(*
SPDX-FileCopyrightText: © 2026 Oleksandr Tiutyk <trofimich@gmail.com>
SPDX-License-Identifier: MIT
License: https://opensource.org/license/mit
*)

(*!
<summary>Provides a scalar natural order for borrowed OBJECT list entries.</summary>
<description>
Supports other ICollectionSortValue objects. Comparisons copy the other scalar key without mutating or
retaining either object. The caller keeps sort keys stable during sorting; no allocation or cleanup is used.
</description>
*)

FUNCTION_BLOCK CollectionComparableProbe EXTENDS TOF_Core.Object IMPLEMENTS ICollectionSortValue
VAR_INPUT
	//! <summary>Scalar key defining the fixture's natural order.</summary>
	SortValue : DINT;
END_VAR
VAR_STAT
	_ClassName : STRING := __POUNAME();
END_VAR

(*!
<summary>Provides the concrete test fixture class name.</summary>
*)
{attribute 'monitoring' := 'call'}
PROPERTY ClassName : REFERENCE TO STRING
GET
ClassName REF= _ClassName;
END_GET
END_PROPERTY

(*!
<summary>Compares supported scalar-key objects and rejects null or unrelated comparable types.</summary>
*)
METHOD CompareTo : TOF_Core.COMPARISON_RESULT
VAR_IN_OUT CONSTANT
	otherValue : TOF_Core.IComparable;
END_VAR
VAR
	otherSortValue : ICollectionSortValue;
	otherKey : DINT;
END_VAR
IF otherValue = 0 THEN
	TOF_Core.Exceptions.ThrowArgumentNotSpecified(
		sourceNamespaceName := NamespaceName,
		sourceClassName := ClassName,
		sourcePOUName := __POUNAME(),
		sourcePosition := __POSITION(),
		argumentName := 'otherValue'
	);
END_IF

IF NOT __QUERYINTERFACE(otherValue, otherSortValue) THEN
	TOF_Core.Exceptions.ThrowStandard(
		sourceNamespaceName := NamespaceName,
		sourceClassName := ClassName,
		sourcePOUName := __POUNAME(),
		sourcePosition := __POSITION(),
		message := "Unsupported collection comparable fixture"
	);
END_IF

otherKey := otherSortValue.GetSortValue();

IF SortValue < otherKey THEN
	CompareTo := TOF_Core.COMPARISON_RESULT.FIRST_LESS_THAN_SECOND;
ELSIF SortValue > otherKey THEN
	CompareTo := TOF_Core.COMPARISON_RESULT.FIRST_GREATER_THAN_SECOND;
ELSE
	CompareTo := TOF_Core.COMPARISON_RESULT.FIRST_EQUAL_TO_SECOND;
END_IF
END_METHOD

(*!
<summary>Copies the configured sort key without mutation.</summary>
*)
METHOD GetSortValue : DINT
GetSortValue := SortValue;
END_METHOD

(*!
<summary>Borrows the compiler-initialized test namespace.</summary>
*)
{attribute 'monitoring' := 'call'}
PROPERTY NamespaceName : REFERENCE TO STRING
GET
NamespaceName REF= CurrentNamespace.Name;
END_GET
END_PROPERTY

(*!
<summary>Reports the complete fixture instance size, excluding separately allocated storage.</summary>
*)
{attribute 'monitoring' := 'call'}
PROPERTY SelfSize : ULINT
GET
SelfSize := XSIZEOF(THIS^);
END_GET
END_PROPERTY

END_FUNCTION_BLOCK

(* stored: Version 1.1.0.1, ProductVersion 3.1.4026.21
   POU CollectionComparableProbe: Id {be1ce13d-533b-447e-b1ca-bc68f369e23c}, SpecialFunc None
   Property ClassName: Id {524c25fa-effd-47d2-899c-109cd5d7359a}
   Get Get: Id {ff64f80e-ffa8-467f-b97b-1226aa0f4865}
   Method CompareTo: Id {ac7bfd62-7bdb-4ae7-a745-a4778e7bded0}
   Method GetSortValue: Id {356150dc-a1f2-4d5a-86ce-b5786a3643b8}
   Property NamespaceName: Id {362a1566-5de6-4e9b-a852-0a7ebe305c75}
   Get Get: Id {b0bab4ca-9949-451d-a46c-f9767d6a89d2}
   Property SelfSize: Id {a9b46d4f-076e-4d4f-9c98-cab3610a380b}
   Get Get: Id {ccbd9b7a-4d0c-4e74-882b-c762762d444a} *)
